// TIA Portal V19 export
// export: Created 2026-10-15T10:10:34.9776652Z, ExportSetting WithDefaults, DisplayName Totally Integrated Automation Portal, DisplayVersion V19, DisplayName TIA Portal Openness, DisplayVersion V19, DisplayName TIA Portal Version Control Interface, DisplayVersion V19, DisplayName STEP 7 Professional, DisplayVersion V19, DisplayName STEP 7 Safety, DisplayVersion V19, DisplayName WinCC Basic/Comfort/Advanced, DisplayVersion V19, DisplayName WinCC Unified, DisplayVersion V19
FUNCTION "ROLL_CounterOp" : Void   // FC8, SCL
{ S7_Optimized_Access := 'TRUE' }
VERSION : 0.1
// stored: AutoNumber true, IsIECCheckEnabled false, SetENOAutomatically false, UDAEnableTagReadback false
   VAR_INPUT
      Number : Int;
      Operation : Int;   // 0=S set; 1=R reset; 2=ZV up; 3=ZR down
      Signal : Bool;
      Preset : Word;
   END_VAR
   VAR_TEMP
      count : Int;
   END_VAR
BEGIN

   IF (#Number < 0) OR (#Number > 127) THEN
       "ROLL_IO".ConversionFault := TRUE;
       RETURN;
   END_IF;
   CASE #Operation OF
       0:
           IF #Signal AND NOT "ROLL_State".S5Counters[#Number].SetPrevious THEN
               #count := "ROLL_DecodeBCD"(Value := #Preset);
               IF #count >= 0 THEN
                   "ROLL_State".S5Counters[#Number].Value := #count;
               END_IF;
           END_IF;
           "ROLL_State".S5Counters[#Number].SetPrevious := #Signal;
       1:
           IF #Signal THEN
               "ROLL_State".S5Counters[#Number].Value := 0;
           END_IF;
       2:
           IF #Signal AND NOT "ROLL_State".S5Counters[#Number].UpPrevious AND ("ROLL_State".S5Counters[#Number].Value < 999) THEN
               "ROLL_State".S5Counters[#Number].Value := "ROLL_State".S5Counters[#Number].Value + 1;
           END_IF;
           "ROLL_State".S5Counters[#Number].UpPrevious := #Signal;
       3:
           IF #Signal AND NOT "ROLL_State".S5Counters[#Number].DownPrevious AND ("ROLL_State".S5Counters[#Number].Value > 0) THEN
               "ROLL_State".S5Counters[#Number].Value := "ROLL_State".S5Counters[#Number].Value - 1;
           END_IF;
           "ROLL_State".S5Counters[#Number].DownPrevious := #Signal;
       ELSE
           "ROLL_IO".ConversionFault := TRUE;
   END_CASE;
END_FUNCTION
